(* IEC 61131-3 sources: JingjiangArm/moonboxpro_arm_8.4/Application/Application/任务列表/LogTask/KS_HY_日志+文件/数据类型+定义, 3 files *)

(* ---- EnumHYLogLevel.st ---- *)
(*@CES
Name=EnumHYLogLevel
Type=Gvl
TypeGuid=2db5746d-d284-4425-9f7f-2663a34b0ebc
Guid=b48dcebc-463e-4092-80ad-422dbcf48ab3
HasDeclaration=True
HasImplementation=False
*)
{DECLARATION}
(*{attribute 'qualified_only'}
{attribute 'strict'}*)
TYPE EnumHYLogLevel :
(
	LOG_LEVEL_INFO	:= 0,(* 一版消息 *)
	LOG_LEVEL_DEBUG	:= 1,(* 调试消息 *)
	LOG_LEVEL_ALARM	:= 2,(* 报警消息 *)
	LOG_LEVEL_ERROR	:= 3,(* 错误消息 *)
	LOG_LEVEL_FATAL	:= 4 (* 严重消息 *)
);
END_TYPE

{IMPLEMENTATION}

(* ---- StHYLogFifo.st ---- *)
(*@CES
Name=StHYLogFifo
Type=Gvl
TypeGuid=2db5746d-d284-4425-9f7f-2663a34b0ebc
Guid=a852f23e-9e5b-4df0-8623-1d9d9541315b
HasDeclaration=True
HasImplementation=False
*)
{DECLARATION}
{attribute 'pack_mode' := '1'}
TYPE StHYLogFifo :
STRUCT
	byIdxR: BYTE;
	byIdxW: BYTE;
	astStHYLogItem: ARRAY [0..255] OF StHYLogItem;
END_STRUCT
END_TYPE

{IMPLEMENTATION}

(* ---- StHYLogItem.st ---- *)
(*@CES
Name=StHYLogItem
Type=Gvl
TypeGuid=2db5746d-d284-4425-9f7f-2663a34b0ebc
Guid=5c0b9e3b-f44a-45e5-a81e-8230d7769e48
HasDeclaration=True
HasImplementation=False
*)
{DECLARATION}
{attribute 'pack_mode' := '1'}
TYPE StHYLogItem :
STRUCT
	sDetails: STRING(200);
END_STRUCT
END_TYPE

{IMPLEMENTATION}
